// TIA Portal V21 export
VAR_GLOBAL   // PLC tag table "TgpUnit_OperandTags"
   TgpUnit_TagFlag AT %M200.0 : Bool;
   TgpUnit_TagTarget AT %M200.1 : Bool;
END_VAR
